// TIA Portal V21 export
// export: Created 2026-11-10T23:32:31.4102164Z, ExportSetting WithDefaults, DisplayName Totally Integrated Automation Portal, DisplayVersion V21 Update 3, DisplayName STEP 7 Professional, DisplayVersion V21 Update 3, DisplayName STEP 7 Safety, DisplayVersion V21, DisplayName Tech WebApplication, DisplayVersion V21, DisplayName WinCC Basic/Comfort/Advanced, DisplayVersion V21 Update 3, DisplayName WinCC Unified, DisplayVersion V21 Update 3
DATA_BLOCK "mTO_InterpreterMapping"   // DB10, Motion_DB
// stored: AutoNumber true, DBAccessibleFromOPCUA true, DBAccessibleFromWebserver true, InstanceOfName TO_InterpreterMapping, OfSystemLibElement TO_InterpreterMapping, OfSystemLibVersion 8.0
TO_InterpreterMapping   // technology object, version 8.0
   // // inherited from TO_Object
BEGIN
END_DATA_BLOCK
